Yaskawa INFORM job: 02025_KOSZ_DO_RURY_70-PLUS-RAMKI.JBI

/JOB
//NAME 02025_KOSZ_DO_RURY_70-PLUS-RAMKI
//POS
///NPOS 218,218,218,0,0,0
///TOOL 0
///POSTYPE PULSE
///PULSE
C00000=-281,-101163,-84214,3730,-80188,-1936
C00001=-281,-101163,-84214,3730,-80188,-1936
C00002=157208,42321,7039,41310,-58295,-11613
C00003=150409,61689,-12910,81671,-34099,-23144
C00004=152528,49836,-26751,84410,-34873,-25218
C00005=152493,38385,-23036,73159,-36698,-18994
C00006=147264,103760,65157,23800,-92258,3726
C00007=146550,104308,54353,23978,-85215,2573
C00008=147295,107763,54133,23856,-83661,2003
C00009=146460,102389,60165,23935,-89859,3533
C00010=145834,34210,-8558,24414,-44224,39072
C00011=144571,58642,-2266,28554,-36050,36909
C00012=145612,62833,-2855,30685,-34156,35502
C00013=144503,52243,3224,24851,-42020,39064
C00014=120555,15135,-34519,-47473,-22108,5770
C00015=123862,59165,-6791,-36652,-28954,-2580
C00016=128755,45321,-19507,-11861,-26051,-11382
C00017=116451,84418,36801,-26901,-79708,-8253
C00018=121869,87599,32734,-28245,-74370,-8901
C00019=120871,90301,31093,-28379,-72550,-8086
C00020=122703,32408,-21346,-21554,-35019,-43815
C00021=130741,49165,-12557,-2398,-28233,-56733
C00022=129681,52067,-14543,-3482,-25555,-55957
C00023=130717,43239,-7941,-2041,-34104,-56920
C00024=126370,89478,49759,-2901,-74617,8364
C00025=130594,106096,57611,-3025,-73915,-173
C00026=135671,99787,49939,-2309,-66778,-1853
C00027=135387,107634,72449,-3249,-82066,-1973
C00028=133977,50927,5217,-3370,-69206,-87684
C00029=131909,54776,-5908,-5184,-49813,-85927
C00030=137525,57587,-2701,-4493,-50055,-88025
C00031=137648,50486,3652,-4076,-57586,-88381
C00032=129358,46579,-1433,-2455,-56315,-83539
C00033=141290,24206,-35414,75400,-30182,-17599
C00034=139321,53340,-22941,89261,-27847,-24192
C00035=140915,41161,-36291,92172,-28651,-26097
C00036=140959,32583,-34967,82519,-29098,-21182
C00037=139136,91856,47671,25542,-85686,5268
C00038=137583,93767,40641,26090,-80431,4664
C00039=138518,97317,39975,26038,-78681,3949
C00040=138336,92285,44735,25767,-83618,5102
C00041=134895,45170,-5214,21800,-38135,42750
C00042=133869,51335,-10602,24985,-31907,41226
C00043=134910,54952,-11675,27339,-29902,39757
C00044=134907,49506,-8526,24066,-34193,41487
C00045=112849,49540,1924,-32526,-41384,-2526
C00046=112828,59759,-6102,-40508,-33092,1964
C00047=112179,46619,-20949,-43189,-31539,3540
C00048=112266,39171,-17616,-37486,-36049,449
C00049=111228,85789,40054,-25860,-82430,-7010
C00050=112245,88973,34515,-26395,-77583,-6282
C00051=111227,92535,34002,-26385,-75941,-5554
C00052=114835,65331,23621,-19065,-65407,-26238
C00053=117108,51630,-11108,-13961,-32795,-44644
C00054=120236,47311,-14449,-6528,-29170,-54657
C00055=119168,50889,-15843,-7919,-26569,-53718
C00056=119453,41895,-10760,-9078,-33755,-50930
C00057=121531,98442,63668,-2340,-81861,2667
C00058=121478,102864,53319,-2407,-73228,2849
C00059=126630,87198,34128,-2212,-59440,1305
C00060=126433,99719,63323,-2678,-80843,1048
C00061=120756,43813,-514,-5728,-59396,-82365
C00062=120756,52460,-8523,-6415,-50076,-81822
C00063=126808,53133,-7797,-5777,-49786,-84038
C00064=126804,46014,-1890,-5265,-57047,-84427
C00065=127789,38302,-24519,78130,-22250,-15987
C00066=127800,48914,-27757,97024,-21678,-25063
C00067=128207,36584,-41501,102088,-22158,-27601
C00068=128383,21926,-38067,77887,-22612,-15996
C00069=129163,87007,35353,27791,-78123,7081
C00070=128167,87997,33431,28141,-76315,6994
C00071=129152,91229,32195,28217,-74464,6189
C00072=128218,83514,39040,27670,-81448,8218
C00073=123752,42492,-9487,16860,-34601,47698
C00074=120103,45558,-16891,7204,-26211,56517
C00075=121114,48915,-18355,8838,-23690,55490
C00076=122605,43213,-10310,16591,-33550,48071
C00077=102322,56250,6520,-35804,-44713,1592
C00078=102282,64934,-18,-41831,-38025,5210
C00079=101000,51872,-15380,-44476,-36504,7022
C00080=100984,42786,-10845,-38470,-42189,3539
C00081=102872,95980,43513,-24260,-81957,-3996
C00082=101975,99505,42873,-24130,-80178,-3328
C00083=102909,93072,46243,-24153,-84865,-4608
C00084=107040,43793,-5997,-15300,-37344,-45079
C00085=108052,49772,-11752,-17509,-30813,-44094
C00086=107092,53578,-12674,-19472,-28594,-42873
C00087=108137,44598,-7832,-15289,-35669,-45300
C00088=112262,101401,62509,-1697,-79856,5796
C00089=112273,105024,56249,-1733,-74145,5871
C00090=117027,94652,43365,-2397,-66509,4438
C00091=117245,99168,60768,-2054,-79818,4138
C00092=109748,45554,2703,-6594,-61258,-78530
C00093=109748,54695,-6001,-7395,-51275,-77872
C00094=115664,53045,-7869,-6899,-50534,-79982
C00095=115664,42198,4108,-5974,-63401,-80755
C00096=114094,42544,4473,10283,-92648,30074
C00097=116764,38974,-24252,19605,-66700,20480
C00098=116764,39826,-24608,19697,-66080,20372
C00099=118338,36457,-17780,18668,-72007,20862
C00100=119061,39982,-23058,19092,-67348,19868
C00101=119061,40795,-23403,19175,-66752,19767
C00102=119061,35980,-20899,18692,-70559,20396
C00103=121044,92533,54944,-1154,-61216,-10928
C00104=124302,166529,126594,-25183,-35107,-49057
C00105=123959,157267,111559,-31709,-30443,-46461
C00106=123959,157736,111044,-32215,-29966,-46201
C00107=123826,155892,108452,-32947,-29465,-45810
C00108=124268,166241,126256,-25250,-35069,-49019
C00109=122293,163687,125144,-26503,-36245,-48217
C00110=119048,153580,110915,-31520,-34220,-45251
C00111=119893,161366,114567,-45012,-31911,-42515
C00112=119893,162037,114301,-45597,-31547,-42207
C00113=119893,162572,123909,-39852,-35758,-45297
C00114=122866,86867,33509,-21111,-15853,-52471
C00115=126243,40965,-18244,-40522,-20964,-50201
C00116=123787,57029,-15218,-60143,-23073,-37730
C00117=123787,57883,-15378,-61258,-22799,-37190
C00118=123664,57468,-15865,-61461,-22817,-37064
C00119=123664,51977,-14480,-54368,-24842,-40523
C00120=123664,51977,-14480,-54368,-24842,-40523
C00121=125295,57830,-13963,-58986,-22538,-38621
C00122=125296,58583,-14115,-59994,-22285,-38134
C00123=125299,50631,-11875,-49840,-25533,-43088
C00124=115650,35746,-12974,33856,-26486,47112
C00125=113547,52477,-17952,29007,-13339,52874
C00126=113547,53192,-18120,30001,-12927,52419
C00127=113692,52974,-18371,30340,-12930,52232
C00128=113692,45275,-15662,21452,-18028,56333
C00129=113692,45275,-15662,21452,-18028,56333
C00130=112101,53810,-15985,25501,-13439,54788
C00131=112049,55073,-16266,26979,-12686,54126
C00132=112025,48327,-14025,19720,-17154,57472
C00133=115359,127852,82120,12682,-35392,60402
C00134=118391,146913,99800,397,-25001,53093
C00135=118391,147433,99318,406,-24437,53089
C00136=118474,146078,97423,534,-23968,53019
C00137=118391,145500,106790,335,-30029,53124
C00138=118451,146260,112190,373,-32961,53102
C00139=118391,145500,106790,335,-30029,53124
C00140=117905,151998,107423,-248,-27081,53456
C00141=117950,152311,106648,-199,-26439,53429
C00142=117887,154325,119178,-226,-33119,53446
C00143=112502,53877,12705,-24757,-100848,-5495
C00144=128780,50425,-557,-26732,-84188,-2205
C00145=131606,47314,-15184,-22938,-73027,-21180
C00146=131854,48845,-16423,-23186,-71538,-20959
C00147=131854,49606,-16698,-23256,-71021,-20854
C00148=131761,49738,-16551,-23228,-71064,-20834
C00149=131854,42444,-13021,-22633,-76515,-21941
C00150=131854,42444,-13021,-22633,-76515,-21941
C00151=132323,50173,-14859,-23280,-71686,-21140
C00152=132434,50775,-15018,-23359,-71283,-21088
C00153=132434,43939,-11435,-22763,-76566,-22139
C00154=138598,52390,-2164,13455,-84086,9906
C00155=104744,-8849,-60671,-33274,-43657,-49146
C00156=92159,-18256,-69173,-34517,-47523,-44903
C00157=91827,4438,-62004,-42729,-49800,-37267
C00158=91818,5680,-62399,-43235,-49147,-36909
C00159=91676,5528,-62533,-43214,-49197,-36874
C00160=91676,5528,-62533,-43214,-49197,-36874
C00161=91827,4438,-62004,-42729,-49800,-37267
C00162=93400,4343,-61853,-42883,-49331,-37711
C00163=93400,5550,-62193,-43369,-48715,-37381
C00164=93167,-5403,-49428,-36047,-58923,-34101
C00165=91827,-17805,-35207,-33276,-72291,-46055
C00166=98842,-11687,-25137,-22009,-69051,-8629
C00167=133516,50989,-3788,-16196,-38937,-20632
C00168=133436,52528,-2466,-16221,-38973,-20603
C00169=133348,52404,-2446,-16230,-39063,-20580
C00170=129075,37367,-6829,-19530,-48616,-16684
C00171=134712,33378,-22556,-16613,-36326,-20658
C00172=129075,37367,-6829,-19530,-48616,-16684
C00173=131059,55248,2023,-20201,-44655,-16677
C00174=130969,57561,3879,-20241,-44632,-16632
C00175=131378,47280,-3853,-19951,-45036,-16909
C00176=127164,32273,-12029,11998,-43670,19984
C00177=121242,44454,-10472,16284,-37844,21983
C00178=121237,46411,-8876,16291,-37822,21980
C00179=121325,46305,-8745,16282,-37967,21967
C00180=124689,31990,-15881,16607,-41417,21066
C00181=124689,31990,-15881,16607,-41417,21066
C00182=124689,31990,-15881,16607,-41417,21066
C00183=122682,44091,-9728,16647,-38725,21464
C00184=122733,44330,-9347,16625,-38838,21466
C00185=122801,45947,-8139,16687,-38770,21420
C00186=122826,31791,-15268,15746,-41548,21965
C00187=125197,9579,-37145,17328,-40006,20532
C00188=115217,-8081,-50354,773,11543,90664
C00189=115990,29069,-9539,-1604,-5188,83946
C00190=118235,28791,-9814,14750,-5334,76366
C00191=117944,18598,-19774,15239,-4422,76186
C00192=138670,25120,-11856,27523,-9237,68458
C00193=139257,34271,-6808,79061,-5026,45511
C00194=137061,32912,-8185,76843,-3549,46783
C00195=137973,21838,-19053,93032,-4042,39448
C00196=137973,21838,-19053,93032,-4042,39448
C00197=137338,33652,-6624,69071,-3913,50209
C00198=135162,32437,-7796,58930,-2552,54999
C00199=135743,24626,-15505,77540,-2624,46642
C00200=110160,22608,-17956,93094,14421,43130
C00201=109051,30359,-10142,96474,15211,41721
C00202=111200,29574,-10921,95955,13756,41674
C00203=110707,19727,-20443,92748,14057,43211
C00204=145779,2561,-42863,153316,-20679,11904
C00205=146612,105798,113888,10829,-72455,18943
C00206=142900,81512,73593,10154,-59860,19165
C00207=142738,84276,76424,10048,-60157,19256
C00208=145684,96477,96590,10823,-66578,18733
C00209=145684,99553,102181,10686,-68407,18902
C00210=145684,99553,102181,10686,-68407,18902
C00211=145315,88062,82572,11036,-62302,18461
C00212=145136,91247,86028,10909,-62761,18573
C00213=145136,100395,103642,10419,-68799,19132
C00214=151636,28907,18690,15103,-54621,14979
C00215=104011,-60420,-74003,22776,-40209,8607
C00216=-281,-101163,-84214,3730,-80188,-1936
C00217=-281,-101163,-84214,3730,-80188,-1936
BC00000=570125
BC00001=299557
BC00002=124171
BC00003=124171
BC00004=124171
BC00005=124171
BC00006=124171
BC00007=124171
BC00008=124171
BC00009=124171
BC00010=124171
BC00011=124171
BC00012=124171
BC00013=124171
BC00014=124171
BC00015=124171
BC00016=124171
BC00017=124171
BC00018=124171
BC00019=124171
BC00020=124171
BC00021=124171
BC00022=124171
BC00023=124171
BC00024=124171
BC00025=124171
BC00026=124171
BC00027=124171
BC00028=124171
BC00029=124171
BC00030=124171
BC00031=124171
BC00032=124171
BC00033=124171
BC00034=124171
BC00035=124171
BC00036=124171
BC00037=124171
BC00038=124171
BC00039=124171
BC00040=124171
BC00041=124171
BC00042=124171
BC00043=124171
BC00044=124171
BC00045=124171
BC00046=124171
BC00047=124171
BC00048=124171
BC00049=124171
BC00050=124171
BC00051=124171
BC00052=124171
BC00053=124171
BC00054=124171
BC00055=124171
BC00056=124171
BC00057=124171
BC00058=124171
BC00059=124171
BC00060=124171
BC00061=124171
BC00062=124171
BC00063=124171
BC00064=124171
BC00065=124171
BC00066=124171
BC00067=124171
BC00068=124171
BC00069=124171
BC00070=124171
BC00071=124171
BC00072=124171
BC00073=124171
BC00074=124171
BC00075=124171
BC00076=124171
BC00077=124171
BC00078=124171
BC00079=124171
BC00080=124171
BC00081=124171
BC00082=124171
BC00083=124171
BC00084=124171
BC00085=124171
BC00086=124171
BC00087=124171
BC00088=124171
BC00089=124171
BC00090=124171
BC00091=124171
BC00092=124171
BC00093=124171
BC00094=124171
BC00095=124171
BC00096=227797
BC00097=227797
BC00098=227797
BC00099=227797
BC00100=352913
BC00101=352913
BC00102=352913
BC00103=227797
BC00104=227797
BC00105=227797
BC00106=227797
BC00107=227797
BC00108=227797
BC00109=227797
BC00110=331582
BC00111=331582
BC00112=331582
BC00113=331582
BC00114=227797
BC00115=227798
BC00116=227798
BC00117=227798
BC00118=227798
BC00119=227798
BC00120=349703
BC00121=349704
BC00122=349704
BC00123=349704
BC00124=227798
BC00125=227798
BC00126=227798
BC00127=227798
BC00128=227798
BC00129=339747
BC00130=339747
BC00131=339747
BC00132=339747
BC00133=227798
BC00134=250331
BC00135=250331
BC00136=250331
BC00137=250331
BC00138=281660
BC00139=363761
BC00140=363761
BC00141=363761
BC00142=363761
BC00143=250331
BC00144=250331
BC00145=250331
BC00146=250331
BC00147=250331
BC00148=250331
BC00149=250331
BC00150=369831
BC00151=369831
BC00152=369831
BC00153=369831
BC00154=250331
BC00155=250331
BC00156=250331
BC00157=250331
BC00158=250331
BC00159=250331
BC00160=250331
BC00161=371627
BC00162=371627
BC00163=371627
BC00164=332143
BC00165=250331
BC00166=250331
BC00167=250331
BC00168=250331
BC00169=250331
BC00170=250331
BC00171=250331
BC00172=363077
BC00173=363077
BC00174=363077
BC00175=363077
BC00176=250331
BC00177=250331
BC00178=250331
BC00179=250331
BC00180=250331
BC00181=250331
BC00182=371513
BC00183=371513
BC00184=371513
BC00185=371513
BC00186=371513
BC00187=250331
BC00188=250331
BC00189=250331
BC00190=250331
BC00191=250331
BC00192=250331
BC00193=250331
BC00194=250331
BC00195=250331
BC00196=360505
BC00197=360505
BC00198=360505
BC00199=360505
BC00200=360505
BC00201=360505
BC00202=360505
BC00203=360505
BC00204=250331
BC00205=250331
BC00206=250331
BC00207=250331
BC00208=250331
BC00209=250331
BC00210=375361
BC00211=375361
BC00212=375361
BC00213=375361
BC00214=250331
BC00215=319701
BC00216=299557
BC00217=570125
EC00000=192,0
EC00001=-931,0
EC00002=-931,0
EC00003=-932,0
EC00004=-932,0
EC00005=-932,0
EC00006=-932,0
EC00007=-932,0
EC00008=-932,0
EC00009=-932,0
EC00010=-932,0
EC00011=-932,0
EC00012=-932,0
EC00013=-932,0
EC00014=-932,0
EC00015=-932,0
EC00016=-932,0
EC00017=-932,0
EC00018=-932,0
EC00019=-932,0
EC00020=-932,0
EC00021=-932,0
EC00022=-932,0
EC00023=-932,0
EC00024=-932,0
EC00025=-932,0
EC00026=-932,0
EC00027=-932,0
EC00028=-932,0
EC00029=-932,0
EC00030=-932,0
EC00031=-932,0
EC00032=-932,0
EC00033=-932,0
EC00034=-932,0
EC00035=-932,0
EC00036=-932,0
EC00037=-932,0
EC00038=-932,0
EC00039=-932,0
EC00040=-932,0
EC00041=-932,0
EC00042=-932,0
EC00043=-932,0
EC00044=-932,0
EC00045=-932,0
EC00046=-932,0
EC00047=-932,0
EC00048=-932,0
EC00049=-932,0
EC00050=-932,0
EC00051=-932,0
EC00052=-932,0
EC00053=-932,0
EC00054=-932,0
EC00055=-932,0
EC00056=-932,0
EC00057=-932,0
EC00058=-932,0
EC00059=-932,0
EC00060=-932,0
EC00061=-932,0
EC00062=-932,0
EC00063=-932,0
EC00064=-932,0
EC00065=-932,0
EC00066=-932,0
EC00067=-932,0
EC00068=-932,0
EC00069=-932,0
EC00070=-932,0
EC00071=-932,0
EC00072=-932,0
EC00073=-932,0
EC00074=-932,0
EC00075=-932,0
EC00076=-932,0
EC00077=-932,0
EC00078=-932,0
EC00079=-932,0
EC00080=-932,0
EC00081=-932,0
EC00082=-933,0
EC00083=-932,0
EC00084=-932,0
EC00085=-932,0
EC00086=-932,0
EC00087=-932,0
EC00088=-932,0
EC00089=-932,0
EC00090=-932,0
EC00091=-932,0
EC00092=-932,0
EC00093=-932,0
EC00094=-933,0
EC00095=-933,0
EC00096=-933,0
EC00097=-933,0
EC00098=-933,0
EC00099=-933,0
EC00100=-933,0
EC00101=-933,0
EC00102=-933,0
EC00103=-933,0
EC00104=-933,0
EC00105=-933,0
EC00106=-933,0
EC00107=-933,0
EC00108=-933,0
EC00109=-933,0
EC00110=-933,0
EC00111=-933,0
EC00112=-933,0
EC00113=-933,0
EC00114=-933,0
EC00115=-933,0
EC00116=-933,0
EC00117=-933,0
EC00118=-933,0
EC00119=-933,0
EC00120=-933,0
EC00121=-933,0
EC00122=-933,0
EC00123=-933,0
EC00124=-933,0
EC00125=-933,0
EC00126=-933,0
EC00127=-933,0
EC00128=-933,0
EC00129=-933,0
EC00130=-933,0
EC00131=-933,0
EC00132=-933,0
EC00133=-933,0
EC00134=-933,0
EC00135=-933,0
EC00136=-933,0
EC00137=-933,0
EC00138=-933,0
EC00139=-933,0
EC00140=-933,0
EC00141=-933,0
EC00142=-933,0
EC00143=-933,0
EC00144=-933,0
EC00145=-933,0
EC00146=-933,0
EC00147=-933,0
EC00148=-933,0
EC00149=-933,0
EC00150=-933,0
EC00151=-933,0
EC00152=-933,0
EC00153=-933,0
EC00154=-933,0
EC00155=-933,0
EC00156=-933,0
EC00157=-933,0
EC00158=-933,0
EC00159=-933,0
EC00160=-933,0
EC00161=-933,0
EC00162=-933,0
EC00163=-933,0
EC00164=38487,0
EC00165=120166,0
EC00166=120166,0
EC00167=120166,0
EC00168=120166,0
EC00169=120166,0
EC00170=120166,0
EC00171=120166,0
EC00172=120166,0
EC00173=120166,0
EC00174=120166,0
EC00175=120166,0
EC00176=120166,0
EC00177=120166,0
EC00178=120166,0
EC00179=120166,0
EC00180=120166,0
EC00181=120166,0
EC00182=120166,0
EC00183=120166,0
EC00184=120166,0
EC00185=120166,0
EC00186=120166,0
EC00187=120166,0
EC00188=120166,0
EC00189=120166,0
EC00190=120166,0
EC00191=120166,0
EC00192=120166,0
EC00193=120166,0
EC00194=120166,0
EC00195=120165,0
EC00196=120165,0
EC00197=120165,0
EC00198=120165,0
EC00199=120165,0
EC00200=120165,0
EC00201=120165,0
EC00202=120165,0
EC00203=120165,0
EC00204=120165,0
EC00205=120165,0
EC00206=120165,0
EC00207=120165,0
EC00208=120165,0
EC00209=120165,0
EC00210=120165,0
EC00211=120165,0
EC00212=120165,0
EC00213=120165,0
EC00214=120165,0
EC00215=-931,0
EC00216=-931,0
EC00217=192,0
//INST
///DATE 2025/05/16 12:39
///ATTR SC,RW
///GROUP1 RB1,BS1
///GROUP2 ST2
NOP
MOVJ C00000 BC00000 VJ=80.00 DEC=20  +MOVJ EC00000 VJ=80.00
MOVJ C00001 BC00001 VJ=80.00 DEC=20  +MOVJ EC00001 VJ=80.00
MOVJ C00002 BC00002 VJ=80.00 DEC=20  +MOVJ EC00002 VJ=80.00
MOVJ C00003 BC00003 VJ=80.00 DEC=20  +MOVJ EC00003 VJ=80.00
MACRO1 MJ#(0) ARGF4
ARCON
WVON WEV#(15)
MOVL C00004 BC00004 V=5.0 DEC=20  +MOVJ EC00004 VJ=80.00
WVOF
ARCOF
MOVJ C00005 BC00005 VJ=80.00 DEC=20  +MOVJ EC00005 VJ=80.00
MOVJ C00006 BC00006 VJ=80.00 DEC=20  +MOVJ EC00006 VJ=80.00
MOVJ C00007 BC00007 VJ=80.00 DEC=20  +MOVJ EC00007 VJ=80.00
ARCON
WVON WEV#(16)
MOVL C00008 BC00008 V=5.0 DEC=20  +MOVJ EC00008 VJ=80.00
WVOF
ARCOF
MOVJ C00009 BC00009 VJ=80.00 DEC=20  +MOVJ EC00009 VJ=80.00
MOVJ C00010 BC00010 VJ=80.00 DEC=20  +MOVJ EC00010 VJ=80.00
MOVJ C00011 BC00011 VJ=80.00 DEC=20  +MOVJ EC00011 VJ=80.00
ARCON
WVON WEV#(16)
MOVL C00012 BC00012 V=5.0 DEC=20  +MOVJ EC00012 VJ=80.00
WVOF
ARCOF
MOVJ C00013 BC00013 VJ=80.00 DEC=20  +MOVJ EC00013 VJ=80.00
MOVJ C00014 BC00014 VJ=80.00 DEC=20  +MOVJ EC00014 VJ=80.00
MOVJ C00015 BC00015 VJ=80.00 DEC=20  +MOVJ EC00015 VJ=80.00
ARCON
WVON WEV#(15)
MOVL C00016 BC00016 V=5.0 DEC=20  +MOVJ EC00016 VJ=80.00
WVOF
ARCOF
MOVJ C00017 BC00017 VJ=80.00 DEC=20  +MOVJ EC00017 VJ=80.00
MOVJ C00018 BC00018 VJ=80.00 DEC=20  +MOVJ EC00018 VJ=80.00
ARCON
WVON WEV#(16)
MOVL C00019 BC00019 V=5.0 DEC=20  +MOVJ EC00019 VJ=80.00
WVOF
ARCOF
MOVJ C00020 BC00020 VJ=80.00 DEC=20  +MOVJ EC00020 VJ=80.00
MOVJ C00021 BC00021 VJ=80.00 DEC=20  +MOVJ EC00021 VJ=80.00
ARCON
WVON WEV#(16)
MOVL C00022 BC00022 V=5.0 DEC=20  +MOVJ EC00022 VJ=80.00
WVOF
ARCOF
MOVJ C00023 BC00023 VJ=80.00 DEC=20  +MOVJ EC00023 VJ=80.00
MOVJ C00024 BC00024 VJ=80.00 DEC=20  +MOVJ EC00024 VJ=80.00
MOVJ C00025 BC00025 VJ=80.00 DEC=20  +MOVJ EC00025 VJ=80.00
ARCON
WVON WEV#(15)
MOVL C00026 BC00026 V=5.0 DEC=20  +MOVJ EC00026 VJ=80.00
WVOF
ARCOF
MOVJ C00027 BC00027 VJ=80.00 DEC=20  +MOVJ EC00027 VJ=80.00
MOVJ C00028 BC00028 VJ=80.00 DEC=20  +MOVJ EC00028 VJ=80.00
MOVJ C00029 BC00029 VJ=80.00 DEC=20  +MOVJ EC00029 VJ=80.00
ARCON
WVON WEV#(15)
MOVL C00030 BC00030 V=5.0 DEC=20  +MOVJ EC00030 VJ=80.00
WVOF
ARCOF
MOVJ C00031 BC00031 VJ=80.00 DEC=20  +MOVJ EC00031 VJ=80.00
MOVJ C00032 BC00032 VJ=80.00 DEC=20  +MOVJ EC00032 VJ=0.78
MOVJ C00033 BC00033 VJ=80.00 DEC=20  +MOVJ EC00033 VJ=0.78
MOVJ C00034 BC00034 VJ=80.00 DEC=20  +MOVJ EC00034 VJ=0.78
ARCON
WVON WEV#(15)
MOVL C00035 BC00035 V=5.0 DEC=20  +MOVJ EC00035 VJ=0.78
WVOF
ARCOF
MOVJ C00036 BC00036 VJ=80.00 DEC=20  +MOVJ EC00036 VJ=80.00
MOVJ C00037 BC00037 VJ=80.00 DEC=20  +MOVJ EC00037 VJ=80.00
MOVJ C00038 BC00038 VJ=80.00 DEC=20  +MOVJ EC00038 VJ=80.00
ARCON
WVON WEV#(16)
MOVL C00039 BC00039 V=5.0 DEC=20  +MOVJ EC00039 VJ=80.00
WVOF
ARCOF
MOVJ C00040 BC00040 VJ=80.00 DEC=20  +MOVJ EC00040 VJ=80.00
MOVJ C00041 BC00041 VJ=80.00 DEC=20  +MOVJ EC00041 VJ=80.00
MOVJ C00042 BC00042 VJ=80.00 DEC=20  +MOVJ EC00042 VJ=80.00
ARCON
WVON WEV#(16)
MOVL C00043 BC00043 V=5.0 DEC=20  +MOVJ EC00043 VJ=80.00
WVOF
ARCOF
MOVJ C00044 BC00044 VJ=80.00 DEC=20  +MOVJ EC00044 VJ=80.00
MOVJ C00045 BC00045 VJ=80.00 DEC=20  +MOVJ EC00045 VJ=80.00
MOVJ C00046 BC00046 VJ=80.00 DEC=20  +MOVJ EC00046 VJ=80.00
ARCON
WVON WEV#(15)
MOVL C00047 BC00047 V=5.0 DEC=20  +MOVJ EC00047 VJ=80.00
WVOF
ARCOF
MOVJ C00048 BC00048 VJ=80.00 DEC=20  +MOVJ EC00048 VJ=80.00
MOVJ C00049 BC00049 VJ=80.00 DEC=20  +MOVJ EC00049 VJ=80.00
MOVJ C00050 BC00050 VJ=80.00 DEC=20  +MOVJ EC00050 VJ=80.00
ARCON
WVON WEV#(16)
MOVL C00051 BC00051 V=5.0 DEC=20  +MOVJ EC00051 VJ=80.00
WVOF
ARCOF
MOVJ C00052 BC00052 VJ=80.00 DEC=20  +MOVJ EC00052 VJ=80.00
MOVJ C00053 BC00053 VJ=80.00 DEC=20  +MOVJ EC00053 VJ=80.00
MOVJ C00054 BC00054 VJ=80.00 DEC=20  +MOVJ EC00054 VJ=80.00
ARCON
WVON WEV#(16)
MOVL C00055 BC00055 V=5.0 DEC=20  +MOVJ EC00055 VJ=80.00
WVOF
ARCOF
MOVJ C00056 BC00056 VJ=80.00 DEC=20  +MOVJ EC00056 VJ=80.00
MOVJ C00057 BC00057 VJ=80.00 DEC=20  +MOVJ EC00057 VJ=80.00
MOVJ C00058 BC00058 VJ=80.00 DEC=20  +MOVJ EC00058 VJ=80.00
ARCON
WVON WEV#(15)
MOVL C00059 BC00059 V=5.0 DEC=20  +MOVJ EC00059 VJ=80.00
WVOF
ARCOF
MOVJ C00060 BC00060 VJ=80.00 DEC=20  +MOVJ EC00060 VJ=80.00
MOVJ C00061 BC00061 VJ=80.00 DEC=20  +MOVJ EC00061 VJ=80.00
MOVJ C00062 BC00062 VJ=80.00 DEC=20  +MOVJ EC00062 VJ=80.00
ARCON
WVON WEV#(15)
MOVL C00063 BC00063 V=5.0 DEC=20  +MOVJ EC00063 VJ=80.00
WVOF
ARCOF
MOVJ C00064 BC00064 VJ=80.00 DEC=20  +MOVJ EC00064 VJ=80.00
MOVJ C00065 BC00065 VJ=30.00 DEC=20  +MOVJ EC00065 VJ=30.00
MOVJ C00066 BC00066 VJ=80.00 DEC=20  +MOVJ EC00066 VJ=80.00
ARCON
WVON WEV#(15)
MOVL C00067 BC00067 V=5.0 DEC=20  +MOVJ EC00067 VJ=80.00
WVOF
ARCOF
MOVJ C00068 BC00068 VJ=80.00 DEC=20  +MOVJ EC00068 VJ=80.00
MOVJ C00069 BC00069 VJ=80.00 DEC=20  +MOVJ EC00069 VJ=80.00
MOVJ C00070 BC00070 VJ=80.00 DEC=20  +MOVJ EC00070 VJ=80.00
ARCON
WVON WEV#(16)
MOVL C00071 BC00071 V=5.0 DEC=20  +MOVJ EC00071 VJ=80.00
WVOF
ARCOF
MOVJ C00072 BC00072 VJ=80.00 DEC=20  +MOVJ EC00072 VJ=80.00
MOVJ C00073 BC00073 VJ=30.00 DEC=20  +MOVJ EC00073 VJ=30.00
MOVJ C00074 BC00074 VJ=80.00 DEC=20  +MOVJ EC00074 VJ=80.00
ARCON
WVON WEV#(16)
MOVL C00075 BC00075 V=5.0 DEC=20  +MOVJ EC00075 VJ=80.00
WVOF
ARCOF
MOVJ C00076 BC00076 VJ=80.00 DEC=20  +MOVJ EC00076 VJ=80.00
MOVJ C00077 BC00077 VJ=80.00 DEC=20  +MOVJ EC00077 VJ=80.00
MOVJ C00078 BC00078 VJ=80.00 DEC=20  +MOVJ EC00078 VJ=80.00
ARCON
WVON WEV#(15)
MOVL C00079 BC00079 V=5.0 DEC=20  +MOVJ EC00079 VJ=80.00
WVOF
ARCOF
MOVJ C00080 BC00080 VJ=80.00 DEC=20  +MOVJ EC00080 VJ=80.00
MOVJ C00081 BC00081 VJ=80.00 DEC=20  +MOVJ EC00081 VJ=80.00
ARCON
WVON WEV#(16)
MOVL C00082 BC00082 V=5.0 DEC=20  +MOVJ EC00082 VJ=80.00
WVOF
ARCOF
MOVJ C00083 BC00083 VJ=80.00 DEC=20  +MOVJ EC00083 VJ=80.00
MOVJ C00084 BC00084 VJ=30.00 DEC=20  +MOVJ EC00084 VJ=30.00
MOVJ C00085 BC00085 VJ=80.00 DEC=20  +MOVJ EC00085 VJ=80.00
ARCON
WVON WEV#(16)
MOVL C00086 BC00086 V=5.0 DEC=20  +MOVJ EC00086 VJ=80.00
WVOF
ARCOF
MOVJ C00087 BC00087 VJ=80.00 DEC=20  +MOVJ EC00087 VJ=80.00
MOVJ C00088 BC00088 VJ=30.00 DEC=20  +MOVJ EC00088 VJ=30.00
MOVJ C00089 BC00089 VJ=30.00 DEC=20  +MOVJ EC00089 VJ=30.00
ARCON
WVON WEV#(15)
MOVL C00090 BC00090 V=5.0 DEC=20  +MOVJ EC00090 VJ=30.00
WVOF
ARCOF
MOVJ C00091 BC00091 VJ=30.00 DEC=20  +MOVJ EC00091 VJ=30.00
MOVJ C00092 BC00092 VJ=30.00 DEC=20  +MOVJ EC00092 VJ=30.00
MOVJ C00093 BC00093 VJ=30.00 DEC=20  +MOVJ EC00093 VJ=30.00
ARCON
WVON WEV#(15)
MOVL C00094 BC00094 V=5.0 DEC=20  +MOVJ EC00094 VJ=30.00
WVOF
ARCOF
MOVJ C00095 BC00095 VJ=80.00 DEC=20  +MOVJ EC00095 VJ=30.00
MOVJ C00096 BC00096 VJ=80.00 DEC=20  +MOVJ EC00096 VJ=0.78
MOVJ C00097 BC00097 VJ=80.00 DEC=20  +MOVJ EC00097 VJ=80.00
MACRO1 MJ#(0) ARGF4
ARCON
WVON WEV#(16)
MOVL C00098 BC00098 V=4.2 DEC=20  +MOVJ EC00098 VJ=80.00
WVOF
ARCOF
MOVJ C00099 BC00099 VJ=80.00 DEC=20  +MOVJ EC00099 VJ=80.00
MOVJ C00100 BC00100 VJ=80.00 DEC=20  +MOVJ EC00100 VJ=50.00
ARCON
MOVL C00101 BC00101 V=4.2 DEC=20  +MOVJ EC00101 VJ=50.00
ARCOF
MOVJ C00102 BC00102 VJ=50.00 DEC=20  +MOVJ EC00102 VJ=50.00
MOVJ C00103 BC00103 VJ=80.00 DEC=20  +MOVJ EC00103 VJ=50.00
MOVJ C00104 BC00104 VJ=80.00 DEC=20  +MOVJ EC00104 VJ=80.00
MOVJ C00105 BC00105 VJ=30.00 DEC=20  +MOVJ EC00105 VJ=80.00
ARCON
WVON WEV#(16)
MOVL C00106 BC00106 V=4.2 DEC=20  +MOVJ EC00106 VJ=80.00
MOVL C00107 BC00107 V=4.2 DEC=20  +MOVJ EC00107 VJ=30.00
WVOF
ARCOF
MOVJ C00108 BC00108 VJ=80.00 DEC=20  +MOVJ EC00108 VJ=80.00
MOVJ C00109 BC00109 VJ=80.00 DEC=20  +MOVJ EC00109 VJ=30.00
MOVJ C00110 BC00110 VJ=80.00 DEC=20  +MOVJ EC00110 VJ=50.00
MOVJ C00111 BC00111 VJ=50.00 DEC=20  +MOVJ EC00111 VJ=50.00
ARCON
WVON WEV#(15)
MOVL C00112 BC00112 V=4.2 DEC=20  +MOVJ EC00112 VJ=50.00
WVOF
ARCOF
MOVJ C00113 BC00113 VJ=80.00 DEC=20  +MOVJ EC00113 VJ=50.00
MOVJ C00114 BC00114 VJ=80.00 DEC=20  +MOVJ EC00114 VJ=30.00
MOVJ C00115 BC00115 VJ=80.00 DEC=20  +MOVJ EC00115 VJ=30.00
MOVJ C00116 BC00116 VJ=80.00 DEC=20  +MOVJ EC00116 VJ=30.00
ARCON
WVON WEV#(16)
MOVL C00117 BC00117 V=4.2 DEC=20  +MOVJ EC00117 VJ=80.00
MOVL C00118 BC00118 V=4.2 DEC=20  +MOVJ EC00118 VJ=80.00
WVOF
ARCOF
MOVJ C00119 BC00119 VJ=80.00 DEC=20  +MOVJ EC00119 VJ=0.78
MOVJ C00120 BC00120 VJ=80.00 DEC=20  +MOVJ EC00120 VJ=50.00
MOVJ C00121 BC00121 VJ=80.00 DEC=20  +MOVJ EC00121 VJ=50.00
ARCON
WVON WEV#(15)
MOVL C00122 BC00122 V=4.2 DEC=20  +MOVJ EC00122 VJ=50.00
WVOF
ARCOF
MOVJ C00123 BC00123 VJ=80.00 DEC=20  +MOVJ EC00123 VJ=50.00
MOVJ C00124 BC00124 VJ=80.00 DEC=20  +MOVJ EC00124 VJ=80.00
MOVJ C00125 BC00125 VJ=80.00 DEC=20  +MOVJ EC00125 VJ=80.00
ARCON
WVON WEV#(16)
MOVL C00126 BC00126 V=4.2 DEC=20  +MOVJ EC00126 VJ=80.00
MOVL C00127 BC00127 V=4.2 DEC=20  +MOVJ EC00127 VJ=80.00
WVOF
ARCOF
MOVJ C00128 BC00128 VJ=80.00 DEC=20  +MOVJ EC00128 VJ=80.00
MOVJ C00129 BC00129 VJ=50.00 DEC=20  +MOVJ EC00129 VJ=50.00
MOVJ C00130 BC00130 VJ=80.00 DEC=20  +MOVJ EC00130 VJ=50.00
ARCON
WVON WEV#(15)
MOVL C00131 BC00131 V=4.2 DEC=20  +MOVJ EC00131 VJ=50.00
WVOF
ARCOF
MOVJ C00132 BC00132 VJ=80.00 DEC=20  +MOVJ EC00132 VJ=50.00
MOVJ C00133 BC00133 VJ=80.00 DEC=20  +MOVJ EC00133 VJ=80.00
MOVJ C00134 BC00134 VJ=80.00 DEC=20  +MOVJ EC00134 VJ=80.00
ARCON
WVON WEV#(16)
MOVL C00135 BC00135 V=4.2 DEC=20  +MOVJ EC00135 VJ=80.00
MOVL C00136 BC00136 V=3.3 DEC=20  +MOVJ EC00136 VJ=80.00
WVOF
ARCOF
MOVJ C00137 BC00137 VJ=50.00 DEC=20  +MOVJ EC00137 VJ=50.00
MOVJ C00138 BC00138 VJ=80.00 DEC=20  +MOVJ EC00138 VJ=80.00
MOVJ C00139 BC00139 VJ=80.00 DEC=20  +MOVJ EC00139 VJ=50.00
MOVJ C00140 BC00140 VJ=80.00 DEC=20  +MOVJ EC00140 VJ=50.00
ARCON
WVON WEV#(15)
MOVL C00141 BC00141 V=4.2 DEC=20  +MOVJ EC00141 VJ=50.00
WVOF
ARCOF
MOVJ C00142 BC00142 VJ=80.00 DEC=20  +MOVJ EC00142 VJ=50.00
MOVJ C00143 BC00143 VJ=80.00 DEC=20  +MOVJ EC00143 VJ=80.00
MOVJ C00144 BC00144 VJ=80.00 DEC=20  +MOVJ EC00144 VJ=80.00
MOVJ C00145 BC00145 VJ=80.00 DEC=20  +MOVJ EC00145 VJ=80.00
MOVJ C00146 BC00146 VJ=80.00 DEC=20  +MOVJ EC00146 VJ=80.00
ARCON
MOVL C00147 BC00147 V=3.3 DEC=20  +MOVJ EC00147 VJ=80.00
MOVL C00148 BC00148 V=3.3 DEC=20  +MOVJ EC00148 VJ=80.00
ARCOF
MOVJ C00149 BC00149 VJ=80.00 DEC=20  +MOVJ EC00149 VJ=80.00
MOVJ C00150 BC00150 VJ=50.00 DEC=20  +MOVJ EC00150 VJ=50.00
MOVJ C00151 BC00151 VJ=50.00 DEC=20  +MOVJ EC00151 VJ=50.00
ARCON
WVON WEV#(15)
MOVL C00152 BC00152 V=4.2 DEC=20  +MOVJ EC00152 VJ=50.00
WVOF
ARCOF
MOVJ C00153 BC00153 VJ=50.00 DEC=20  +MOVJ EC00153 VJ=50.00
MOVJ C00154 BC00154 VJ=80.00 DEC=20  +MOVJ EC00154 VJ=80.00
MOVJ C00155 BC00155 VJ=80.00 DEC=20  +MOVJ EC00155 VJ=80.00
MOVJ C00156 BC00156 VJ=80.00 DEC=20  +MOVJ EC00156 VJ=80.00
MOVJ C00157 BC00157 VJ=80.00 DEC=20  +MOVJ EC00157 VJ=80.00
ARCON
WVON WEV#(15)
MOVL C00158 BC00158 V=4.2 DEC=20  +MOVJ EC00158 VJ=80.00
MOVL C00159 BC00159 V=4.2 DEC=20  +MOVJ EC00159 VJ=80.00
WVOF
ARCOF
MOVJ C00160 BC00160 VJ=50.00 DEC=20  +MOVJ EC00160 VJ=50.00
MOVJ C00161 BC00161 VJ=50.00 DEC=20  +MOVJ EC00161 VJ=50.00
MOVJ C00162 BC00162 VJ=50.00 DEC=20  +MOVJ EC00162 VJ=50.00
ARCON
WVON WEV#(15)
MOVL C00163 BC00163 V=4.2 DEC=20  +MOVJ EC00163 VJ=50.00
WVOF
ARCOF
MOVJ C00164 BC00164 VJ=50.00 DEC=20  +MOVJ EC00164 VJ=50.00
MOVJ C00165 BC00165 VJ=80.00 DEC=20  +MOVJ EC00165 VJ=80.00
MOVJ C00166 BC00166 VJ=80.00 DEC=20  +MOVJ EC00166 VJ=80.00
MOVJ C00167 BC00167 VJ=80.00 DEC=20  +MOVJ EC00167 VJ=80.00
ARCON
WVON WEV#(15)
MOVL C00168 BC00168 V=4.2 DEC=20  +MOVJ EC00168 VJ=80.00
WVOF
MOVJ C00169 BC00169 VJ=80.00 DEC=20  +MOVJ EC00169 VJ=80.00
ARCOF
MOVJ C00170 BC00170 VJ=80.00 DEC=20  +MOVJ EC00170 VJ=80.00
MOVJ C00171 BC00171 VJ=50.00 DEC=20  +MOVJ EC00171 VJ=50.00
MOVJ C00172 BC00172 VJ=50.00 DEC=20  +MOVJ EC00172 VJ=50.00
MOVJ C00173 BC00173 VJ=50.00 DEC=20  +MOVJ EC00173 VJ=50.00
ARCON
WVON WEV#(15)
MOVL C00174 BC00174 V=4.2 DEC=20  +MOVJ EC00174 VJ=50.00
WVOF
ARCOF
MOVJ C00175 BC00175 VJ=50.00 DEC=20  +MOVJ EC00175 VJ=50.00
MOVJ C00176 BC00176 VJ=80.00 DEC=20  +MOVJ EC00176 VJ=80.00
MOVJ C00177 BC00177 VJ=80.00 DEC=20  +MOVJ EC00177 VJ=80.00
ARCON
WVON WEV#(15)
MOVL C00178 BC00178 V=4.2 DEC=20  +MOVJ EC00178 VJ=80.00
WVOF
MOVL C00179 BC00179 V=3.3 DEC=20  +MOVJ EC00179 VJ=80.00
ARCOF
MOVJ C00180 BC00180 VJ=80.00 DEC=20  +MOVJ EC00180 VJ=80.00
MOVJ C00181 BC00181 VJ=50.00 DEC=20  +MOVJ EC00181 VJ=50.00
MOVJ C00182 BC00182 VJ=50.00 DEC=20  +MOVJ EC00182 VJ=50.00
MOVJ C00183 BC00183 VJ=50.00 DEC=20  +MOVJ EC00183 VJ=50.00
MOVJ C00184 BC00184 VJ=50.00 DEC=20  +MOVJ EC00184 VJ=50.00
ARCON
WVON WEV#(15)
MOVL C00185 BC00185 V=4.2 DEC=20  +MOVJ EC00185 VJ=50.00
WVOF
ARCOF
MOVJ C00186 BC00186 VJ=50.00 DEC=20  +MOVJ EC00186 VJ=50.00
MOVJ C00187 BC00187 VJ=80.00 DEC=20  +MOVJ EC00187 VJ=80.00
MOVJ C00188 BC00188 VJ=80.00 DEC=20  +MOVJ EC00188 VJ=80.00
MOVJ C00189 BC00189 VJ=80.00 DEC=20  +MOVJ EC00189 VJ=80.00
ARCON
MOVL C00190 BC00190 V=5.0 DEC=20  +MOVJ EC00190 VJ=80.00
ARCOF
MOVJ C00191 BC00191 VJ=10.00 DEC=20  +MOVJ EC00191 VJ=80.00
MOVJ C00192 BC00192 VJ=10.00 DEC=20  +MOVJ EC00192 VJ=10.00
MOVJ C00193 BC00193 VJ=10.00 DEC=20  +MOVJ EC00193 VJ=10.00
ARCON
MOVL C00194 BC00194 V=5.0 DEC=20  +MOVJ EC00194 VJ=10.00
ARCOF
MOVJ C00195 BC00195 VJ=10.00 DEC=20  +MOVJ EC00195 VJ=10.00
MOVJ C00196 BC00196 VJ=80.00 DEC=20  +MOVJ EC00196 VJ=50.00
MOVJ C00197 BC00197 VJ=80.00 DEC=20  +MOVJ EC00197 VJ=80.00
ARCON
MOVL C00198 BC00198 V=4.2 DEC=20  +MOVJ EC00198 VJ=80.00
ARCOF
MOVJ C00199 BC00199 VJ=80.00 DEC=20  +MOVJ EC00199 VJ=80.00
MOVJ C00200 BC00200 VJ=80.00 DEC=20  +MOVJ EC00200 VJ=80.00
MOVJ C00201 BC00201 VJ=80.00 DEC=20  +MOVJ EC00201 VJ=80.00
ARCON
MOVL C00202 BC00202 V=4.2 DEC=20  +MOVJ EC00202 VJ=80.00
ARCOF
MOVJ C00203 BC00203 VJ=80.00 DEC=20  +MOVJ EC00203 VJ=80.00
MOVJ C00204 BC00204 VJ=10.00 DEC=20  +MOVJ EC00204 VJ=10.00
MOVJ C00205 BC00205 VJ=10.00 DEC=20  +MOVJ EC00205 VJ=10.00
MOVJ C00206 BC00206 VJ=10.00 DEC=20  +MOVJ EC00206 VJ=10.00
ARCON
WVON WEV#(15)
MOVL C00207 BC00207 V=4.2 DEC=20  +MOVJ EC00207 VJ=10.00
WVOF
ARCOF
MOVJ C00208 BC00208 VJ=80.00 DEC=20  +MOVJ EC00208 VJ=10.00
MOVJ C00209 BC00209 VJ=80.00 DEC=20  +MOVJ EC00209 VJ=80.00
MOVJ C00210 BC00210 VJ=80.00 DEC=20  +MOVJ EC00210 VJ=80.00
MOVJ C00211 BC00211 VJ=80.00 DEC=20  +MOVJ EC00211 VJ=80.00
ARCON
WVON WEV#(15)
MOVL C00212 BC00212 V=4.2 DEC=20  +MOVJ EC00212 VJ=80.00
WVOF
ARCOF
MOVJ C00213 BC00213 VJ=80.00 DEC=20  +MOVJ EC00213 VJ=80.00
MOVJ C00214 BC00214 VJ=50.00 DEC=20  +MOVJ EC00214 VJ=10.00
MOVJ C00215 BC00215 VJ=50.00 DEC=20  +MOVJ EC00215 VJ=50.00
MOVJ C00216 BC00216 VJ=80.00 DEC=20  +MOVJ EC00216 VJ=80.00
MOVJ C00217 BC00217 VJ=80.00 DEC=20  +MOVJ EC00217 VJ=80.00
END
